Staubli VAL3: _productCycle.pgx

public program _productCycle()
  local bool l_bErr
  local bool l_bStartClock
  local num l_nClock
  local num l_nLastAct
  local num l_nLibIndex
  local string l_sPath
begin
  //do
  // rs:nPLCcmd=0
  //等待数据库切换完成以及程序号完成
  // wait(io:dInput[30]==true)
  //wait(bBool==true)
  //
  waitEndMove()
  //
  //（工作号&程序号->切换完成->plc启动信号->productcycle->（工作号&程序号->切换完成->plc启动信号
  //
  //获取程序号
  call io:getAnaIO(io:aInItem[0].aAio,rs:nProgCode,l_bErr)
  switch rs:nProgCode
    case 0
      //call prog:makeTraj("test")
    break
    case 1
      rs:sTrajStatus="开始执行prod01"
      call prog:makeTraj("prod01")

    break
    case 2
      rs:sTrajStatus="开始执行prod02"
      call prog:makeTraj("prod02")

    break
    case 3
      rs:sTrajStatus="开始执行prod03"
      call prog:makeTraj("prod03")

    break
    case 4
      rs:sTrajStatus="开始执行prod04"
      call prog:makeTraj("prod04")

    break
    case 5
      rs:sTrajStatus="开始执行prod05"
      call prog:makeTraj("prod05")

    break
    case 6
      rs:sTrajStatus="开始执行prod06"
      call prog:makeTraj("prod06")

    break
    case 7
      rs:sTrajStatus="开始执行prod07"
      call prog:makeTraj("prod07")

    break
    case 8
      rs:sTrajStatus="开始执行prod08"
      call prog:makeTraj("prod08")

    break
    case 9
      rs:sTrajStatus="开始执行prod09"
      call prog:makeTraj("prod09")

    break
    case 10
      rs:sTrajStatus="开始执行prod10"
      call prog:makeTraj("prod10")

    break
    case 11
      rs:sTrajStatus="开始执行prod11"
      call prog:makeTraj("prod11")

    break
    case 12
      rs:sTrajStatus="开始执行prod012"
      call prog:makeTraj("prod12")

    break
    case 13
      rs:sTrajStatus="开始执行prod13"
      call prog:makeTraj("prod13")

    break
    case 14
      rs:sTrajStatus="开始执行prod14"
      call prog:makeTraj("prod14")

    break
    case 15
      rs:sTrajStatus="开始执行prod15"
      call prog:makeTraj("prod15")

    break
    case 16
      rs:sTrajStatus="开始执行prod16"
      call prog:makeTraj("prod16")

    break


    case 17
      rs:sTrajStatus="开始执行prod17"
      call prog:makeTraj("prod17")
    break

    case 18
      rs:sTrajStatus="开始执行prod18"
      call prog:makeTraj("prod18")
    break
    case 19
      rs:sTrajStatus="开始执行prod19"
      call prog:makeTraj("prod19")
    break

    case 20
      rs:sTrajStatus="开始执行prod20"
      call prog:makeTraj("prod20")
    break

    case 21
      rs:sTrajStatus="开始执行prod21"
      call prog:makeTraj("prod21")

    break
    case 22
      rs:sTrajStatus="开始执行prod22"
      call prog:makeTraj("prod22")

    break
    case 23
      rs:sTrajStatus="开始执行prod23"
      call prog:makeTraj("prod23")

    break
    case 24
      rs:sTrajStatus="开始执行prod24"
      call prog:makeTraj("prod24")

    break
    case 25
      rs:sTrajStatus="开始执行prod25"
      call prog:makeTraj("prod25")

    break
    case 26
      rs:sTrajStatus="开始执行prod26"
      call prog:makeTraj("prod26")

    break
    case 27
      rs:sTrajStatus="开始执行prod27"
      call prog:makeTraj("prod27")

    break
    case 28
      rs:sTrajStatus="开始执行prod28"
      call prog:makeTraj("prod28")

    break
    case 29
      rs:sTrajStatus="开始执行prod29"
      call prog:makeTraj("prod29")

    break
    case 30
      rs:sTrajStatus="开始执行prod30"
      call prog:makeTraj("prod30")

    break
    case 31
      rs:sTrajStatus="开始执行prod31"
      call prog:makeTraj("prod31")

    break
    case 32
      rs:sTrajStatus="开始执行prod032"
      call prog:makeTraj("prod32")

    break
    case 33
      rs:sTrajStatus="开始执行prod33"
      call prog:makeTraj("prod33")

    break
    case 34
      rs:sTrajStatus="开始执行prod34"
      call prog:makeTraj("prod34")

    break
    case 35
      rs:sTrajStatus="开始执行prod35"
      call prog:makeTraj("prod35")

    break
    case 36
      rs:sTrajStatus="开始执行prod36"
      call prog:makeTraj("prod36")

    break

    case 37
      rs:sTrajStatus="开始执行prod37"
      call prog:makeTraj("prod37")
    break

    case 38
      rs:sTrajStatus="开始执行prod38"
      call prog:makeTraj("prod38")
    break
    case 39
      rs:sTrajStatus="开始执行prod39"
      call prog:makeTraj("prod39")
    break

    case 40
      rs:sTrajStatus="开始执行prod40"
      call prog:makeTraj("prod40")
    break
    case 40
      rs:sTrajStatus="开始执行prod40"
      call prog:makeTraj("prod40")

    break
    case 41
      rs:sTrajStatus="开始执行prod41"
      call prog:makeTraj("prod41")

    break
    case 42
      rs:sTrajStatus="开始执行prod042"
      call prog:makeTraj("prod42")

    break
    case 43
      rs:sTrajStatus="开始执行prod43"
      call prog:makeTraj("prod43")

    break
    case 44
      rs:sTrajStatus="开始执行prod44"
      call prog:makeTraj("prod44")

    break
    case 45
      rs:sTrajStatus="开始执行prod45"
      call prog:makeTraj("prod45")

    break
    case 46
      rs:sTrajStatus="开始执行prod46"
      call prog:makeTraj("prod46")

    break

    case 47
      rs:sTrajStatus="开始执行prod47"
      call prog:makeTraj("prod47")
    break

    case 48
      rs:sTrajStatus="开始执行prod48"
      call prog:makeTraj("prod48")
    break
    case 49
      rs:sTrajStatus="开始执行prod49"
      call prog:makeTraj("prod49")
    break

    case 50
      rs:sTrajStatus="开始执行prod50"
      call prog:makeTraj("prod50")
    break

  endSwitch
  if l_bStartClock and l_nLastAct!=rs:nActCode
    rs:_nCTIndex=(rs:_nCTIndex+1)%size(rs:_nCycleTime)
    rs:_nCycleTime[rs:_nCTIndex]=clock()-l_nClock
  else
    l_bStartClock=true
  endIf
  l_nClock=clock()
  l_nLastAct=rs:nActCode
  //delay(0)
  //
  rs:_nOmacStat=1
  rs:sTrajStatus=""
  rs:_sRobotStatus="当前件生产结束"
  //2025.1.6 add 结束扭矩记录程序
  if taskStatus("getForce")!=-1
    delay(0.2)
    taskKill("getForce")
  endIf
end
